(* IEC 61131-3 sources: Claude/ballplate-sim/codesys, 2 files *)

(* ---- FB_BallCtrl.st ---- *)
// Function block FB_BallCtrl : one axis of the ball-and-plate controller.
// Plant is (almost) a double integrator:  x'' = (5/7) * g * theta
// so a PD law with the 5/7*g gain scaled out gives chosen wn / zeta:
//     theta = ( wn^2 * (sp - x) - 2*zeta*wn * (v_hat - sp_vel) ) / k
// Same algorithm as CascadePD in ballplate/mock_plc.py (which is tested against the simulator).
FUNCTION_BLOCK FB_BallCtrl
VAR_INPUT
    bEnable     : BOOL;
    rSetpoint   : REAL;                 // m
    rSetpointVel: REAL;                 // m/s velocity feed-forward (0 for fixed setpoint)
    rPos        : REAL;                 // m, measured
    rDt         : REAL := 0.01;         // s, task cycle time (use the task interval!)
    rWn         : REAL := 1.5;          // rad/s  closed-loop natural frequency
    rZeta       : REAL := 0.9;
    rVelTau     : REAL := 0.06;         // s, velocity filter time constant
    rKi         : REAL := 0.15;         // integral gain (fights rolling resistance)
    rMaxDeg     : REAL := 10.0;
END_VAR
VAR_OUTPUT
    rTiltCmdDeg : REAL;                 // deg
END_VAR
VAR
    rPosPrev    : REAL;
    rVel        : REAL;
    rInteg      : REAL;                 // rad
    bInit       : BOOL;
    rErr, rCmd, rA : REAL;
END_VAR
VAR CONSTANT
    K_PLANT     : REAL := 7.0071;       // 5/7 * 9.81
    RAD2DEG     : REAL := 57.29578;
END_VAR

IF NOT bEnable THEN
    rInteg := 0; bInit := FALSE; rTiltCmdDeg := 0; RETURN;
END_IF
IF NOT bInit THEN rPosPrev := rPos; rVel := 0; bInit := TRUE; END_IF

// filtered derivative of the measured position
rA := rDt / (rVelTau + rDt);
rVel := rVel + rA * ((rPos - rPosPrev) / rDt - rVel);
rPosPrev := rPos;

rErr := rSetpoint - rPos;
rInteg := LIMIT(-0.05, rInteg + rKi * rErr * rDt, 0.05);
rCmd := (rWn*rWn*rErr - 2.0*rZeta*rWn*(rVel - rSetpointVel)) / K_PLANT + rInteg;
rTiltCmdDeg := LIMIT(-rMaxDeg, rCmd * RAD2DEG, rMaxDeg);

(* ---- PLC_PRG_Example.st ---- *)
// Example PLC program for the rolling-table simulator (task interval 10 ms).
// Uses the IO words from the project's GVL "gIo":
//   outputs  F_YR10, F_YR20 : INT   tilt X / Y   (+-32000 <-> +-15 deg)
//   inputs   F_XG12, F_XG22 : INT   distance X/Y (+-32000 <-> +-1 m)
//            F_XG11, F_XG21 : INT   velocity X/Y (-32000..+32000 <-> vel_min..vel_max, default +-0.4 m/s)
//            F_XG10, F_XG20 : INT   acceleration (+-32000 <-> +-9.81 m/s^2)
// The ranges must match [scaling] in config/sim.toml of the simulator.
PROGRAM PLC_PRG_Example
VAR
    fbX, fbY    : FB_BallCtrl;
    bRun        : BOOL := TRUE;
    rSpX, rSpY  : REAL;                  // m, ball setpoint (0,0 = centre)
    rPosX, rPosY: REAL;                  // m, scaled measurements
    rTiltX, rTiltY : REAL;               // deg, controller outputs
END_VAR

// raw -> engineering units
rPosX := -1.0 + (INT_TO_REAL(gIo.F_XG12) + 32000.0) / 64000.0 * 2.0;
rPosY := -1.0 + (INT_TO_REAL(gIo.F_XG22) + 32000.0) / 64000.0 * 2.0;

fbX(bEnable := bRun, rSetpoint := rSpX, rSetpointVel := 0.0, rPos := rPosX, rDt := 0.01);
fbY(bEnable := bRun, rSetpoint := rSpY, rSetpointVel := 0.0, rPos := rPosY, rDt := 0.01);
rTiltX := fbX.rTiltCmdDeg;
rTiltY := fbY.rTiltCmdDeg;

// engineering units -> raw (limited to the INT range)
gIo.F_YR10 := REAL_TO_INT(LIMIT(-32000.0, rTiltX / 15.0 * 32000.0, 32000.0));
gIo.F_YR20 := REAL_TO_INT(LIMIT(-32000.0, rTiltY / 15.0 * 32000.0, 32000.0));
